(*
SPDX-FileCopyrightText: © 2026 Oleksandr Tiutyk <trofimich@gmail.com>
SPDX-License-Identifier: MIT
License: https://opensource.org/license/mit
*)

(*!
<summary>Provides fluent assertions on a copied DINT value.</summary>
<description>
Copies actual into persistent instance storage before the entry method returns; literals and expression
results therefore remain valid throughout the immediate chain. Owns no heap allocation or pointed-to resource.
The message prefixes every failure until the next preparation. Finish one chain before starting another on
the owning Assertions provider. Use only from the owning test callback on one task, without reentry.
Obtain this context from the owning provider; direct unprepared use is unsupported.
Expected arguments use the declared IEC type; ordinary compiler conversions happen before comparison.
This context does not depend on another assertion context.
Object metadata is available before preparation; inherited equality compares instance identity.
</description>
*)

{attribute 'no_explicit_call' := 'do not call this function block directly'}
FUNCTION_BLOCK DIntAssertionContext EXTENDS TOF_Core.Object
VAR_STAT
	{attribute 'hide'}
	_ClassName : STRING := __POUNAME();
END_VAR
VAR
	_Actual : DINT;
	_TestCase : ITestCase;
	_Message : WSTRING(255);
END_VAR

(*!
<summary>Provides the implementation class name.</summary>
<description>
Borrowed read-only reference to compiler-initialized storage, valid throughout the instance lifetime.
Do not modify the returned reference; no ownership is transferred.
</description>
*)
{attribute 'monitoring' := 'call'}
PROPERTY ClassName : REFERENCE TO STRING
GET
ClassName REF= _ClassName;
END_GET
END_PROPERTY

(*!
<summary>Asserts that the actual value is strictly greater than expected.</summary>
<description>
Records failure without interrupting the callback; preserves the message for the rest of the chain.
</description>
<param name="expected">Expected value converted by the compiler to DINT.</param>
*)
METHOD FINAL IsGreaterThan : REFERENCE TO DIntAssertionContext
VAR_INPUT
	expected : DINT;
END_VAR
IF _Actual <= expected THEN
	failComparison(
		expected := expected,
		expectation := "Expected value > "
	);
END_IF

IsGreaterThan REF= THIS^;
END_METHOD

(*!
<summary>Asserts that the actual value meets the inclusive lower boundary.</summary>
<description>
Records failure without interrupting the callback; preserves the message for the rest of the chain.
</description>
<param name="expected">Expected value converted by the compiler to DINT.</param>
*)
METHOD FINAL IsGreaterThanOrEquals : REFERENCE TO DIntAssertionContext
VAR_INPUT
	expected : DINT;
END_VAR
IF _Actual < expected THEN
	failComparison(
		expected := expected,
		expectation := "Expected value >= "
	);
END_IF

IsGreaterThanOrEquals REF= THIS^;
END_METHOD

(*!
<summary>Asserts that the actual value is strictly less than expected.</summary>
<description>
Records failure without interrupting the callback; preserves the message for the rest of the chain.
</description>
<param name="expected">Expected value converted by the compiler to DINT.</param>
*)
METHOD FINAL IsLessThan : REFERENCE TO DIntAssertionContext
VAR_INPUT
	expected : DINT;
END_VAR
IF _Actual >= expected THEN
	failComparison(
		expected := expected,
		expectation := "Expected value < "
	);
END_IF

IsLessThan REF= THIS^;
END_METHOD

(*!
<summary>Asserts that the actual value meets the inclusive upper boundary.</summary>
<description>
Records failure without interrupting the callback; preserves the message for the rest of the chain.
</description>
<param name="expected">Expected value converted by the compiler to DINT.</param>
*)
METHOD FINAL IsLessThanOrEquals : REFERENCE TO DIntAssertionContext
VAR_INPUT
	expected : DINT;
END_VAR
IF _Actual > expected THEN
	failComparison(
		expected := expected,
		expectation := "Expected value <= "
	);
END_IF

IsLessThanOrEquals REF= THIS^;
END_METHOD

(*!
<summary>Provides the library namespace.</summary>
<description>
Borrowed read-only reference to the compiler-initialized namespace, valid throughout the instance lifetime.
Do not modify the returned reference; no ownership is transferred.
</description>
*)
{attribute 'monitoring' := 'call'}
PROPERTY NamespaceName : REFERENCE TO STRING
GET
NamespaceName REF= CurrentNamespace.Name;
END_GET
END_PROPERTY

(*!
<summary>Asserts inequality with the expected value.</summary>
<description>
Records failure without interrupting the callback; preserves the message for the rest of the chain.
</description>
<param name="expected">Expected value converted by the compiler to DINT.</param>
*)
METHOD FINAL NotToBe : REFERENCE TO DIntAssertionContext
VAR_INPUT
	expected : DINT;
END_VAR
IF _Actual = expected THEN
	failComparison(
		expected := expected,
		expectation := "Expected value not to be: "
	);
END_IF

NotToBe REF= THIS^;
END_METHOD

(*!
<summary>Copies the actual operand and replaces the chain-wide message.</summary>
<description>
Called by the owning Assertions provider after it verifies the running test case.
No pointer to this method's input storage is retained. The receiver is borrowed until the next preparation;
the owning provider keeps it alive throughout the immediate chain.
</description>
<param name="actual">Value copied into this context.</param>
<param name="testCase">Borrowed failure receiver for the immediate chain.</param>
<param name="message">Copied diagnostic prefix, including empty to clear the previous prefix.</param>
*)
METHOD INTERNAL FINAL Prepare
VAR_INPUT
	actual : DINT;
	testCase : ITestCase;
	message : WSTRING(255);
END_VAR
_Actual := actual;
_TestCase := testCase;
_Message := message;
END_METHOD

(*!
<summary>Reports the byte size of this concrete instance.</summary>
<description>
Includes inline fields and nested instances, but excludes separately allocated payloads.
Obtaining the size does not transfer ownership or validate an arbitrary address.
</description>
*)
{attribute 'monitoring' := 'call'}
PROPERTY SelfSize : ULINT
GET
SelfSize := XSIZEOF(THIS^);
END_GET
END_PROPERTY

(*!
<summary>Asserts equality with the expected value.</summary>
<description>
Records failure without interrupting the callback; preserves the message for the rest of the chain.
</description>
<param name="expected">Expected value converted by the compiler to DINT.</param>
*)
METHOD FINAL ToBe : REFERENCE TO DIntAssertionContext
VAR_INPUT
	expected : DINT;
END_VAR
IF _Actual <> expected THEN
	failComparison(
		expected := expected,
		expectation := "Expected: "
	);
END_IF

ToBe REF= THIS^;
END_METHOD

(*!
<summary>Formats a failed typed predicate and reports it with the chain message.</summary>
<description>
Does not change operands or chain state. The receiver retains its first failure. Reporting exceptions
propagate to the enclosing test callback handler; an unprepared receiver is a configuration error.
</description>
<param name="expected">Typed expected operand used only for this diagnostic.</param>
<param name="expectation">Prefix identifying the failed predicate.</param>
*)
METHOD PRIVATE failComparison
VAR_INPUT
	expected : DINT;
	expectation : WSTRING(40);
END_VAR
VAR
	actualText : WSTRING(255);
	expectedText : WSTRING(255);
	diagnostic : TOF_Core.ERROR_MESSAGE;
END_VAR
actualText := TO_WSTRING(_Actual);
expectedText := TO_WSTRING(expected);

diagnostic := TOF_Core.WideStrings.Concat255(
	expectation,
	expectedText,
	", but was: ",
	actualText
);

TestServices.ReportAssertionFailure(
	testCase := _TestCase,
	message := _Message,
	sourceClassName := ClassName,
	defaultMessage := diagnostic
);
END_METHOD

END_FUNCTION_BLOCK

(* stored: Version 1.1.0.1
   POU DIntAssertionContext: Id {be53c725-cf41-45f3-a0e9-b7a462c934b3}, SpecialFunc None
   Folder Service methods: Id {38841bb8-741b-4496-9075-e42ec5b29ab2}
   Property ClassName: Id {daf68f08-b054-4367-b5b1-a9ea38a7d604}
   Get Get: Id {8a275ac6-4172-468a-b419-eb90d757ddf5}
   Method IsGreaterThan: Id {940f4b25-ac00-43f5-8297-347cfbcd80cf}
   Method IsGreaterThanOrEquals: Id {6acb8268-d454-4efa-bba8-9e10b3d60319}
   Method IsLessThan: Id {3c6a30e6-808d-4690-a0b3-cbb227764d1a}
   Method IsLessThanOrEquals: Id {3281e4af-2a67-45cc-973c-8e911b205fed}
   Property NamespaceName: Id {989d47f9-e303-4562-b417-bbbf03834778}
   Get Get: Id {5811234b-e832-4ea2-8735-66de04065548}
   Method NotToBe: Id {00ad172d-00fe-4e12-a880-06aa54689b2b}
   Method Prepare: Id {4de53826-db87-41d0-a3e6-1ccaf1168d6e}
   Property SelfSize: Id {6f8b12b5-e391-434e-8db8-4422588a7996}
   Get Get: Id {2aa8f44c-6c40-477f-8550-7849f4e85784}
   Method ToBe: Id {bb9ba507-c693-45dd-a2ad-c037aff8fb45}
   Method failComparison: Id {58420bef-7ba4-43b3-915f-6bdbc925ae18} *)
